Fanuc KAREL source: kt00038.KL

-- PROVISIONAL review KL for V940-1; original PC SHA256 9facd4450cf3087773b290f6fdbf51b17fc02acc22e6d9a116f9a98ed9761c77
-- Incomplete behavior may be omitted. Consult companion uncertainty JSON. Do not deploy.
PROGRAM KT00038
%NOLOCKGROUP
VAR
  I1 : INTEGER
  OUT : REAL
-- UNRESOLVED_DECL Y2 type=002018
BEGIN
  -- V9_ZERO_TABLE_METADATA_HINT layout=0001; no indexed target words; source/name/runtime held
  -- UNRESOLVED_PC offsets 5-16; opcodes 2E,23
  -- UNRESOLVED_PC offsets 21-35; opcodes 2E,22,9D,33,B2
  -- UNRESOLVED_PC offsets 40-63; opcodes 21,22,9D,33,B1,53,64,23
  -- UNRESOLVED_PC offsets 68-72; opcodes 7F
END KT00038
